(* IEC 61131-3 sources: POMIRTS_lab3/AS/Library_2/AsHydCon/V3.10.0 (part 2) *)

(* ---- AsHydCon.fun ---- *)
(********************************************************************
 * COPYRIGHT -- B&R
 ********************************************************************
 * Library: AsHydCon
 * File: AsHydCon.fun
 * Author: DI Thomas J. Frauscher
 * Created: July 2011
 ********************************************************************
 * Function blocks of library AsHydCon
 ********************************************************************)

FUNCTION_BLOCK HCRPT1 (*1st order delay element.*)
	VAR_INPUT
		enable : BOOL; (*Enable function block.*)
		V : REAL; (*Gain. Units: [1].*)
		T1 : REAL; (*Time constant. Units: [s]. Valid value range: T1 >= 0.*)
		u : REAL; (*Input value.*)
		Set_y : USINT; (*"Apply preset value for y" controller input. Valid value range: {0,1,2}.*)
		y_set : REAL; (*Preset value for y.*)
	END_VAR
	VAR_OUTPUT
		y : REAL; (*Output value.*)
		status : UINT; (*Function block status message.*)
	END_VAR
	VAR
		Internal : HCRPT1_Internal_typ; (*Data for internal use.*)
	END_VAR
END_FUNCTION_BLOCK

FUNCTION_BLOCK HCRPT2 (*2nd order delay element.*)
	VAR_INPUT
		enable : BOOL; (*Enable function block.*)
		V : REAL; (*Gain. Units: [1].*)
		T1 : REAL; (*Time constant 1. Units: [s]. Valid value range: T1 >= 0.*)
		T2 : REAL; (*Time constant 2. Units: [s]. Valid value range: T2 >= 0.*)
		u : REAL; (*Input value.*)
		Set_y : USINT; (*"Apply preset value for y" controller input. Valid value range: {0,1,2}.*)
		y_set : REAL; (*Preset value for y.*)
	END_VAR
	VAR_OUTPUT
		y : REAL; (*Output value.*)
		status : UINT; (*Function block status message.*)
	END_VAR
	VAR
		Internal : HCRPT2_Internal_typ; (*Data for internal use.*)
	END_VAR
END_FUNCTION_BLOCK

FUNCTION_BLOCK HCRPT2s (*Oscillating 2nd order delay element.*)
	VAR_INPUT
		enable : BOOL; (*Enable function block.*)
		V : REAL; (*Gain. Units: [1].*)
		D : REAL; (*Damping constant. Units: [1]. Valid value range: D >= 0.*)
		Tf : REAL; (*Filter time constant. Units: [s]. Valid value range: Tf > 0.*)
		u : REAL; (*Input value.*)
		Set_y : USINT; (*"Apply preset value for y" controller input. Valid value range: {0,1,2}.*)
		y_set : REAL; (*Preset value for y.*)
	END_VAR
	VAR_OUTPUT
		y : REAL; (*Output value.*)
		status : UINT; (*Function block status message.*)
	END_VAR
	VAR
		Internal : HCRPT2s_Internal_typ; (*Data for internal use.*)
	END_VAR
END_FUNCTION_BLOCK

FUNCTION_BLOCK HCRDT1 (*1st order differentiator.*)
	VAR_INPUT
		enable : BOOL; (*Enable function block.*)
		Tv : REAL; (*Differentiation time constant. Units: [s]. Valid value range: Tv >= 0.*)
		Tf : REAL; (*Filter time constant. Units: [s]. Valid value range: Tf >= 0.*)
		u : REAL; (*Input value.*)
		n_Avg : USINT; (*Moving average filter for the input value u. Valid value range: {0, 1, 2, ..., 100}.*)
		Reset_y : USINT; (*Reset controller input y to 0. Valid value range: {0,1,2}.*)
	END_VAR
	VAR_OUTPUT
		y : REAL; (*Output value.*)
		status : UINT; (*Function block status message.*)
	END_VAR
	VAR
		Internal : HCRDT1_Internal_typ; (*Data for internal use.*)
	END_VAR
END_FUNCTION_BLOCK

FUNCTION_BLOCK HCRDT2 (*2nd order differentiator.*)
	VAR_INPUT
		enable : BOOL; (*Enable function block.*)
		Tv : REAL; (*Differentiation time constant. Units: [s]. Valid value range: Tv >= 0.*)
		T1 : REAL; (*Filter time constant 1. Units: [s]. Valid value range: T1 >= 0.*)
		T2 : REAL; (*Filter time constant 2. Units: [s]. Valid value range: T2 >= 0.*)
		u : REAL; (*Input value.*)
		n_Avg : USINT; (*Moving average filter for the input value u. Valid value range: {0, 1, 2, ..., 100}.*)
		Reset_y : USINT; (*Reset controller input y to 0. Valid value range: {0,1,2}.*)
	END_VAR
	VAR_OUTPUT
		y : REAL; (*Output value.*)
		status : UINT; (*Function block status message.*)
	END_VAR
	VAR
		Internal : HCRDT2_Internal_typ; (*Data for internal use.*)
	END_VAR
END_FUNCTION_BLOCK

FUNCTION_BLOCK HCRDT2s (*Oscillating 2nd order differentiator.*)
	VAR_INPUT
		enable : BOOL; (*Enable function block.*)
		D : REAL; (*Damping constant. Units: [1]. Valid value range: D >= 0.*)
		Tv : REAL; (*Differentiation time constant. Units: [s]. Valid value range: Tv >= 0.*)
		Tf : REAL; (*Filter time constant. Units: [s]. Valid value range: Tf >= 0.*)
		u : REAL; (*Input value.*)
		Reset_y : USINT; (*Reset controller input y to 0. Valid value range: {0,1,2}.*)
	END_VAR
	VAR_OUTPUT
		y : REAL; (*Output value.*)
		status : UINT; (*Function block status message.*)
	END_VAR
	VAR
		Internal : HCRDT2s_Internal_typ; (*Data for internal use.*)
	END_VAR
END_FUNCTION_BLOCK

FUNCTION_BLOCK HCRIT1 (*1st order integrator.*)
	VAR_INPUT
		enable : BOOL; (*Enable function block.*)
		V : REAL; (*Gain. Units: [1].*)
		Tn : REAL; (*Integration time constant (integral action time). Units: [s]. Valid value range: Tn > 0.*)
		T1 : REAL; (*Time constant. Units: [s]. Valid value range: T1 >= 0.*)
		u : REAL; (*Input value.*)
		Set_y : USINT; (*"Apply preset value for y" controller input. Valid value range: {0,1,2}.*)
		y_set : REAL; (*Preset value for y.*)
	END_VAR
	VAR_OUTPUT
		y : REAL; (*Output value.*)
		status : UINT; (*Function block status message.*)
	END_VAR
	VAR
		Internal : HCRIT1_Internal_typ; (*Data for internal use.*)
	END_VAR
END_FUNCTION_BLOCK

FUNCTION_BLOCK HCRNotch (*2nd order notch filter.*)
	VAR_INPUT
		enable : BOOL; (*Enable function block.*)
		V : REAL; (*Gain. Units: [1].*)
		f0 : REAL; (*Filter frequency. Units: [Hz]. Valid value range: f0 > 0.*)
		B : REAL; (*Filter band width. Units: [Hz]. Valid value range: B > 0.*)
		u : REAL; (*Input value.*)
		Set_y : USINT; (*"Apply preset value for y" controller input. Valid value range: {0,1,2}.*)
		y_set : REAL; (*Preset value for y.*)
	END_VAR
	VAR_OUTPUT
		y : REAL; (*Output value.*)
		status : UINT; (*Function block status message.*)
	END_VAR
	VAR
		Internal : HCRNotch_Internal_typ; (*Data for internal use.*)
	END_VAR
END_FUNCTION_BLOCK

FUNCTION_BLOCK HCRPT1cP (*Converging 1st order delay element.*)
	VAR_INPUT
		enable : BOOL; (*Enable function block.*)
		T1 : REAL; (*Time constant. Units: [s]. Valid value range: T1 >= 0.*)
		u : REAL; (*Input value.*)
		Set_y : USINT; (*"Apply preset value for y" controller input. Valid value range: {0,1,2}.*)
		y_set : REAL; (*Preset value for y.*)
	END_VAR
	VAR_OUTPUT
		y : REAL; (*Output value.*)
		status : UINT; (*Function block status message.*)
	END_VAR
	VAR
		Internal : HCRPT1cP_Internal_typ; (*Data for internal use.*)
	END_VAR
END_FUNCTION_BLOCK

FUNCTION_BLOCK HCRJoltFree (*Jolt-free switching between 2 inputs.*)
	VAR_INPUT
		enable : BOOL; (*Enable function block.*)
		tSwitch : REAL; (*Switching time. Units: [s]. Valid value range: tSwitch >= 0.*)
		uSwitch : BOOL; (*Switch between signal inputs u1 and u2.*)
		u1 : REAL; (*Input value 1.*)
		u2 : REAL; (*Input value 2.*)
	END_VAR
	VAR_OUTPUT
		y : REAL; (*Output value.*)
		status : UINT; (*Function block status message.*)
	END_VAR
	VAR
		Internal : HCRJoltFree_Internal_typ; (*Data for internal use.*)
		PT1cP : HCRPT1cP; (*Internally used function block.*)
	END_VAR
END_FUNCTION_BLOCK

FUNCTION_BLOCK HCRFIFO (*FIFO (dead time) element.*)
	VAR_INPUT
		enable : BOOL; (*Enable function block.*)
		t_FIFO : DINT; (*Delay time. Units: [µs].*)
		x : REAL; (*Input value.*)
		Set_y : BOOL; (*"Apply preset value for y" controller input.*)
		y_set : REAL; (*Preset value for y.*)
	END_VAR
	VAR_OUTPUT
		y : REAL; (*Output value.*)
		status : UINT; (*Function block status message.*)
	END_VAR
	VAR
		Internal : HCRFIFO_Internal_typ; (*Data for internal use.*)
	END_VAR
END_FUNCTION_BLOCK

FUNCTION_BLOCK HCRRampGen (*Ramp generator.*)
	VAR_INPUT
		enable : BOOL; (*Enable function block.*)
		t_rise : REAL; (*Rise time. Units [s]. Valid value range: t_rise >= 0.*)
		t_hold : REAL; (*Constant holding time. Units [s]. Valid value range: t_hold >= 0.*)
		t_fall : REAL; (*Fall time. Units [s]. Valid value range: t_fall >= 0.*)
		y_start : REAL; (*Start value for the output value y.*)
		y_hold : REAL; (*Stop value for the output value y.*)
		y_end : REAL; (*End value for the output value y.*)
		Init : BOOL; (*Based on the start value y_start, Init = 1 initiates a new ramp that ends with an end value y_end, after crossing a stop phase t_hold with stop value y_hold.*)
	END_VAR
	VAR_OUTPUT
		y : REAL; (*Ramp generator output value.*)
		dy : REAL; (*Time derivative (dy/dt) of y.*)
		dy_ramped : REAL; (*Ramped time derivative (dy/dt) of y.*)
		Finished : BOOL; (*Finished = 1 indicates the end of ramp generation.*)
		status : UINT; (*Function block status message.*)
	END_VAR
	VAR
		Internal : HCRRampGen_Internal_typ; (*Data for internal use.*)
	END_VAR
END_FUNCTION_BLOCK

FUNCTION_BLOCK HCRSPF (*Smart path finder.*)
	VAR_INPUT
		enable : BOOL; (*Enable function block.*)
		pMove_Para : REFERENCE TO HCRMovePara_typ; (*Movement parameters (t_Jolt, vC_pos, vC_neg, aAcc_pos, aDec_pos, aAcc_neg, aDec_neg).*)
		Stop : BOOL; (*Stop = 1 stops trajectory planning.*)
		s_home : REAL; (*Homing position. Units: [mm].*)
		Set_home : BOOL; (*If no set trajectory is being processed at the moment, setting Set_home = 1 sets s_set = s_home and Reached = 1.*)
		s_end : REAL; (*End position of the trajectory. Units: [mm].*)
		Init : BOOL; (*Based on the current set position s_set and the current set speed v_set, Init = 1 initiates a new trajectory that ends at the point s_end.*)
		Brake : BOOL; (*Based on the current values of s_set and v_set, Brake = 1 stops the movement with the delay aDec_pos (positive direction) or aDec_neg (negative direction).*)
	END_VAR
	VAR_OUTPUT
		s_set : REAL; (*Set position. Units: [mm].*)
		v_set : REAL; (*Set speed. Units: [mm/s]. Value range: -vC_neg <= v_set <= vC_pos.*)
		a_set : REAL; (*Set acceleration. Units: [mm/s²]. Value range: -max(aDec_pos, aDec_neg) <= a_set <= max(aAcc_pos, aAcc_neg).*)
		MoveDir : SINT; (*Direction of movement. Value range: {-3,-2,-1: negative direction of movement (-3: Deceleration phase, -2: Constant speed phase, -1: Acceleration phase), 0: standstill, 1,2,3: positive direction of movement (1: Acceleration phase, 2: Constant speed phase, 3: Deceleration phase)}.*)
		ApproachDir : SINT; (*Approach direction indicates in which direction the end position s_end is reached. Value range: {-1: negative approach direction, 0: undefined, 1: positive approach direction}.*)
		Reached : BOOL; (*Reached = 1 indicates that the end position has been reached and that the movement is complete.*)
		status : UINT; (*Function block status message.*)
	END_VAR
	VAR
		Internal : HCRSPF_Internal_typ; (*Data for internal use.*)
		SystemInfo : SysInfo; (*Internally used function block.*)
	END_VAR
END_FUNCTION_BLOCK

FUNCTION_BLOCK HCRSFG (*Smart force generator.*)
	VAR_INPUT
		enable : BOOL; (*Enable function block.*)
		t_Jolt : REAL; (*Jolt time. Units [s]. Valid value range: 0 <= t_Jolt <= 0.2.*)
		Stop : BOOL; (*Stop = 1 stops trajectory planning.*)
		dFp_home : REAL; (*Homing value for the set force rate. Units: [N/s].*)
		Fp_home : REAL; (*Homing value for the set force. Units: [N].*)
		Set_home : BOOL; (*If no set trajectory is being processed at the moment, setting Set_home = 1 sets Fp_set = Fp_home, dFp_set = dFp_home and Reached = 1.*)
		t_delta : REAL; (*Time difference specified for bringing Fp_set from its present value to the end value Fp_end. Units: [s]. Valid value range: t_delta > t_Jolt.*)
		Fp_end : REAL; (*End value of the set force trajectory. Units: [N].*)
		Init : BOOL; (*Based on the current set force Fp_set and the current set force rate dFp_set, Init = 1 initiates a new trajectory that ends at the point Fp_end (dFp_set = 0).*)
	END_VAR
	VAR_OUTPUT
		Fp_set : REAL; (*Set force. Units: [N].*)
		dFp_set : REAL; (*Set force rate. Units: [N/s].*)
		t_delta_act : REAL; (*Actual time difference needed for bringing Fp_set to the specified end value Fp_end. Units: [s]. Value range: t_delta_act > t_Jolt.*)
		Reached : BOOL; (*Reached = 1 indicates that end value of the set force has been reached and that the profile generation is complete.*)
		status : UINT; (*Function block status message.*)
	END_VAR
	VAR
		Internal : HCRSFG_Internal_typ; (*Data for internal use.*)
		SPF : HCRSPF; (*Internally used function block.*)
	END_VAR
END_FUNCTION_BLOCK

FUNCTION_BLOCK HCRAutoTune (*Autotuning-algorithm for Kp.*)
	VAR_INPUT
		enable : BOOL; (*Enable function block.*)
		pSupply_max : REAL; (*Maximum system pressure (supply pressure). Units: [bar]. Valid value range: pSupply_max >= 0.*)
		A_Cyl_pos : REAL; (*Cylinder piston area whose pressurization induces a movement in the positive direction (e.g. extending piston). Units: [cm]. Valid value range: A_Cyl_pos > 0.*)
		A_Cyl_neg : REAL; (*Cylinder piston area whose pressurization induces a movement in the negative direction (e.g. retracting piston). Units: [cm]. Valid value range: A_Cyl_neg > 0.*)
		Qnom_pos : REAL; (*Nominal valve-volume flow, which, together with A_Cyl_pos results in a movement in the positive direction (e.g. extending piston). Units: [l/min]. Valid value range: Qnom_pos > 0.*)
		Qnom_neg : REAL; (*Nominal valve-volume flow, which, together with A_Cyl_neg results in a movement in the negative direction (e.g. retracting piston). Units: [l/min]. Valid value range: Qnom_neg > 0.*)
		pDelta_nom : REAL; (*Nominal pressure drop at valve edge. Units: [bar]. Valid value range: pDelta_nom > 0.*)
		V0_pos : REAL; (*Static volume in reference to the cylinder chamber responsible for movement in the 'positive' direction (e.g. extending piston). Units: [l]. Valid value range: V0_pos >= 0.*)
		V0_neg : REAL; (*Static volume in reference to the cylinder chamber responsible for movement in the 'negative' direction (e.g. retracting piston). Units: [l]. Valid value range: V0_neg >= 0.*)
		h_Cyl : REAL; (*Cylinder height. Units: [mm]. Valid value range: h_Cyl > 0.*)
		m_Cyl : REAL; (*Resulting mass of the moving hydraulic system. Units: [kg]. Valid value range: m_Cyl > 0.*)
		s_min : REAL; (*Minimum value of set position and actual position. Units: [mm]. Valid value range: s_min < s_max.*)
		s_max : REAL; (*Maximum value of set position and actual position. Units: [mm]. Valid value range: s_max > s_min.*)
		Update : USINT; (*Any changes to the above variables (pSupply_max, A_Cyl_pos, ..., s_max) must be applied with Update = 1.*)
	END_VAR
	VAR_OUTPUT
		Kp : REAL; (*Calculated proportional gain of the position controller. Units: [1].*)
		status : UINT; (*Function block status message.*)
	END_VAR
	VAR
		Internal : HCRAutoTune_Internal_typ; (*Data for internal use.*)
	END_VAR
END_FUNCTION_BLOCK

FUNCTION_BLOCK HCROmega0 (*Omega0-correction for Kp.*)
	VAR_INPUT
		enable : BOOL; (*Enable function block.*)
		A_Cyl_pos : REAL; (*Cylinder piston area whose pressurization induces a movement in the positive direction (e.g. extending piston). Units: [cm]. Valid value range: A_Cyl_pos > 0.*)
		A_Cyl_neg : REAL; (*Cylinder piston area whose pressurization induces a movement in the negative direction (e.g. retracting piston). Units: [cm]. Valid value range: A_Cyl_neg > 0.*)
		V0_pos : REAL; (*Static volume in reference to the cylinder chamber responsible for movement in the 'positive' direction (e.g. extending piston). Units: [l]. Valid value range: V0_pos >= 0.*)
		V0_neg : REAL; (*Static volume in reference to the cylinder chamber responsible for movement in the 'negative' direction (e.g. retracting piston). Units: [l]. Valid value range: V0_neg >= 0.*)
		h_Cyl : REAL; (*Cylinder height. Units: [mm]. Valid value range: h_Cyl > 0.*)
		x_Cyl_min : REAL; (*Minimum value of x_Cyl until a correction of the proportional gain of the position controller has been calculated. Units: [mm]. Valid value range: 0 <= x_Cyl_min < x_Cyl_max.*)
		x_Cyl_max : REAL; (*Maximum value of x_Cyl until a correction of the proportional gain of the position controller has been calculated. Units: [mm]. Valid value range: x_Cyl_min < x_Cyl_max <= h_Cyl.*)
		Update : USINT; (*Any changes to the above variables (A_Cyl_pos, A_Cyl_neg, ..., x_Cyl_max) must be applied with Update = 1.*)
		x_Cyl : REAL; (*Current position of the cylinder piston (always based on the cylinder). Units: [mm]. Valid value range: 0 <= x_Cyl <= h_Cyl.*)
	END_VAR
	VAR_OUTPUT
		x0_Cyl : REAL; (*Position of cylinder piston at which the critical natural frequency of the hydraulic system occurs. Units: [mm]. Value range: 0 <= x0_Cyl <= h_Cyl.*)
		Kp_xCorr : REAL; (*Calculated multiplication factor for correcting the proportional gain of the position controller with Kp_xCorr = Kp_xCorr(x_Cyl). Units: [1]. Value range: 1 <= Kp_xCorr <= 2.*)
		status : UINT; (*Function block status message.*)
	END_VAR
	VAR
		Internal : HCROmega0_Internal_typ; (*Data for internal use.*)
	END_VAR
END_FUNCTION_BLOCK

FUNCTION_BLOCK HCRvyServo (*v-y servo correction (pressure).*)
	VAR_INPUT
		enable : BOOL; (*Enable function block.*)
		pSupply_max : REAL; (*Maximum system pressure (supply pressure). Units: [bar]. Valid value range: pSupply_max >= 0.*)
		pSupply : REAL; (*System pressure (supply pressure). Units: [bar]. Valid value range: pSupply > 0.*)
		pTank : REAL; (*Tank pressure. Units: [bar]. Valid value range: pTank >= 0.*)
		A_Cyl_pos : REAL; (*Cylinder piston area whose pressurization induces a movement in the positive direction (e.g. extending piston). Units: [cm]. Valid value range: A_Cyl_pos > 0.*)
		A_Cyl_neg : REAL; (*Cylinder piston area whose pressurization induces a movement in the negative direction (e.g. retracting piston). Units: [cm]. Valid value range: A_Cyl_neg > 0.*)
		Qnom_pos : REAL; (*Nominal valve-volume flow, which, together with A_Cyl_pos results in a movement in the positive direction (e.g. extending piston). Units: [l/min]. Valid value range: Qnom_pos > 0.*)
		Qnom_neg : REAL; (*Nominal valve-volume flow, which, together with A_Cyl_neg results in a movement in the negative direction (e.g. retracting piston). Units: [l/min]. Valid value range: Qnom_neg > 0.*)
		pDelta_nom : REAL; (*Nominal pressure drop at valve edge. Units: [bar]. Valid value range: pDelta_nom > 0.*)
		yValve_0 : REAL; (*Valve overlap. Units: [1]. Valid value range:  0 <= yValve_0 < 1.*)
		yValve_min : REAL; (*Minimum valve opening (|yValve| = yValve_min). Units: [1]. Valid value range: 0 <= yValve_min <= 1.*)
		Neg_y : BOOL; (*Negative values for the valve opening yValve result in a positive speed, and vice versa (inverted valve behavior).*)
		Update : USINT; (*Any changes to the above variables must be applied with Update = (Mode + 1).*)
		pCyl_pos : REAL; (*Chamber pressure for movement in the 'positive' direction. Units: [bar]. Valid value range: 0 <= pCyl_pos < pSupply.*)
		pCyl_neg : REAL; (*Chamber pressure for movement in the 'negative' direction. Units: [bar]. Valid value range: 0 <= pCyl_neg < pSupply.*)
		vCyl_abs : REAL; (*Absolute speed of cylinder movement. Units: [mm/s]. Valid value range: -vCyl_sup < vCyl_abs < vCyl_sup.*)
		vCyl_rel : REAL; (*Relative speed of cylinder movement. Units: [%]. Valid value range: -100 <= vCyl_rel <= 100.*)
		Zero_yValve : BOOL; (*Setting this input results in the immediate output of yValve = 0 and Qy = 0.*)
	END_VAR
	VAR_OUTPUT
		Qy_abs : REAL; (*Volume flow produced by vCyl_abs (Qy = Qy_abs + Qy_rel). Units: [l/min]. Value range: -Qnom_neg <= Qy_abs <= Qnom_pos.*)
		Qy_rel : REAL; (*Volume flow produced by vCyl_rel (Qy_rel = Qy - Qy_abs). Units: [l/min]. Value range: -Qnom_neg <= Qy_rel <= Qnom_pos.*)
		Qy : REAL; (*Volume flow produced by valve opening yValve. Units: [l/min]. Value range: -Qnom_neg <= Qy <= Qnom_pos.*)
		yValve : REAL; (*Valve opening. Units: [1]. Value range: -1 <= yValve <= 1.*)
		MoveDir : SINT; (*Direction of movement. Value range: {-1: negative direction of movement, 0: undefined, 1: positive direction of movement}.*)
		status : UINT; (*Function block status message.*)
	END_VAR
	VAR
		Internal : HCRvyServo_Internal_typ; (*Data for internal use.*)
	END_VAR
END_FUNCTION_BLOCK

FUNCTION_BLOCK HCRvyServo_Fp (*v-y servo correction (force).*)
	VAR_INPUT
		enable : BOOL; (*Enable function block.*)
		pSupply_max : REAL; (*Maximum system pressure (supply pressure). Units: [bar]. Valid value range: pSupply_max >= 0.*)
		pSupply : REAL; (*System pressure (supply pressure). Units: [bar]. Valid value range: pSupply > 0.*)
		pTank : REAL; (*Tank pressure. Units: [bar]. Valid value range: pTank >= 0.*)
		A_Cyl_pos : REAL; (*Cylinder piston area whose pressurization induces a movement in the positive direction (e.g. extending piston). Units: [cm]. Valid value range: A_Cyl_pos > 0.*)
		A_Cyl_neg : REAL; (*Cylinder piston area whose pressurization induces a movement in the negative direction (e.g. retracting piston). Units: [cm]. Valid value range: A_Cyl_neg > 0.*)
		Qnom_pos : REAL; (*Nominal valve-volume flow, which, together with A_Cyl_pos results in a movement in the positive direction (e.g. extending piston). Units: [l/min]. Valid value range: Qnom_pos > 0.*)
		Qnom_neg : REAL; (*Nominal valve-volume flow, which, together with A_Cyl_neg results in a movement in the negative direction (e.g. retracting piston). Units: [l/min]. Valid value range: Qnom_neg > 0.*)
		pDelta_nom : REAL; (*Nominal pressure drop at valve edge. Units: [bar]. Valid value range: pDelta_nom > 0.*)
		yValve_0 : REAL; (*Valve overlap. Units: [1]. Valid value range:  0 <= yValve_0 < 1.*)
		yValve_min : REAL; (*Minimum valve opening (|yValve| = yValve_min). Units: [1]. Valid value range: 0 <= yValve_min <= 1.*)
		Neg_y : BOOL; (*Negative values for the valve opening yValve result in a positive speed, and vice versa (inverted valve behavior).*)
		Update : USINT; (*Any changes to the above variables must be applied with Update = (Mode + 1).*)
		Fp_Cyl : REAL; (*Process force. Units: [N].*)
		Ff_Cyl_pos : REAL; (*Friction force in positive direction. Units: [N]. Valid value range:  Ff_Cyl_pos >= 0.*)
		Ff_Cyl_neg : REAL; (*Friction force in negative direction. Units: [N]. Valid value range:  Ff_Cyl_neg >= 0.*)
		vCyl_abs : REAL; (*Absolute speed of cylinder movement. Units: [mm/s]. Valid value range: -vCyl_sup < vCyl_abs < vCyl_sup.*)
		vCyl_rel : REAL; (*Relative speed of cylinder movement. Units: [%]. Valid value range: -100 <= vCyl_rel <= 100.*)
		Zero_yValve : BOOL; (*Setting this input results in the immediate output of yValve = 0 and Qy = 0.*)
	END_VAR
	VAR_OUTPUT
		Qy_abs : REAL; (*Volume flow produced by vCyl_abs (Qy = Qy_abs + Qy_rel). Units: [l/min]. Value range: -Qnom_neg <= Qy_abs <= Qnom_pos.*)
		Qy_rel : REAL; (*Volume flow produced by vCyl_rel (Qy_rel = Qy - Qy_abs). Units: [l/min]. Value range: -Qnom_neg <= Qy_rel <= Qnom_pos.*)
		Qy : REAL; (*Volume flow produced by valve opening yValve. Units: [l/min]. Value range: -Qnom_neg <= Qy <= Qnom_pos.*)
		yValve : REAL; (*Valve opening. Units: [1]. Value range: -1 <= yValve <= 1.*)
		MoveDir : SINT; (*Direction of movement. Value range: {-1: negative direction of movement, 0: undefined, 1: positive direction of movement}.*)
		status : UINT; (*Function block status message.*)
	END_VAR
	VAR
		Internal : HCRvyServo_Fp_Internal_typ; (*Data for internal use.*)
	END_VAR
END_FUNCTION_BLOCK

FUNCTION_BLOCK HCRFyServo (*F-y servo correction (pressure).*)
	VAR_INPUT
		enable : BOOL; (*Enable function block.*)
		pSupply_max : REAL; (*Maximum system pressure (supply pressure). Units: [bar]. Valid value range: pSupply_max >= 0.*)
		pSupply : REAL; (*System pressure (supply pressure). Units: [bar]. Valid value range: pSupply > 0.*)
		pTank : REAL; (*Tank pressure. Units: [bar]. Valid value range: pTank >= 0.*)
		A_Cyl_pos : REAL; (*Cylinder piston area whose pressurization induces a movement in the positive direction (e.g. extending piston). Units: [cm]. Valid value range: A_Cyl_pos > 0.*)
		A_Cyl_neg : REAL; (*Cylinder piston area whose pressurization induces a movement in the negative direction (e.g. retracting piston). Units: [cm]. Valid value range: A_Cyl_neg > 0.*)
		Qnom_pos : REAL; (*Nominal valve-volume flow, which, together with A_Cyl_pos results in a movement in the positive direction (e.g. extending piston). Units: [l/min]. Valid value range: Qnom_pos > 0.*)
		Qnom_neg : REAL; (*Nominal valve-volume flow, which, together with A_Cyl_neg results in a movement in the negative direction (e.g. retracting piston). Units: [l/min]. Valid value range: Qnom_neg > 0.*)
		pDelta_nom : REAL; (*Nominal pressure drop at valve edge. Units: [bar]. Valid value range: pDelta_nom > 0.*)
		yValve_0 : REAL; (*Valve overlap. Units: [1]. Valid value range:  0 <= yValve_0 < 1.*)
		V0_pos : REAL; (*Static volume in reference to the cylinder chamber responsible for movement in the 'positive' direction (e.g. extending piston). Units: [l]. Valid value range: V0_pos >= 0.*)
		V0_neg : REAL; (*Static volume in reference to the cylinder chamber responsible for movement in the 'negative' direction (e.g. retracting piston). Units: [l]. Valid value range: V0_neg >= 0.*)
		h_Cyl : REAL; (*Cylinder height. Units: [mm]. Valid value range: h_Cyl > 0.*)
		Neg_y : BOOL; (*Negative values for the valve opening yValve result in a positive speed, and vice versa (inverted valve behavior).*)
		Update : USINT; (*Any changes to the above variables must be applied with Update = (Mode + 1).*)
		x_Cyl : REAL; (*Current position of the cylinder piston (always based on the cylinder). Units: [mm]. Valid value range: 0 <= x_Cyl <= h_Cyl.*)
		v_Cyl : REAL; (*Current speed of the cylinder piston (always based on the cylinder). Units: [mm].*)
		pCyl_pos : REAL; (*Chamber pressure for movement in the 'positive' direction. Units: [bar]. Valid value range: 0 <= pCyl_pos < pSupply.*)
		pCyl_neg : REAL; (*Chamber pressure for movement in the 'negative' direction. Units: [bar]. Valid value range: 0 <= pCyl_neg < pSupply.*)
		dF_Cyl_abs : REAL; (*Absolute rate of force increase of the cylinder. Units: [N/s]. Valid value range:  -dF_Cyl_sup < dF_Cyl_abs < dF_Cyl_sup.*)
		dF_Cyl_rel : REAL; (*Relative rate of force increase of the cylinder. Units: [%]. Valid value range: -100 <= dF_Cyl_rel <= 100.*)
	END_VAR
	VAR_OUTPUT
		Qy : REAL; (*Volume flow produced by valve opening yValve. Units: [l/min]. Value range: -Qnom_neg <= Qy <= Qnom_pos.*)
		yValve : REAL; (*Valve opening. Units: [1]. Value range: -1 <= yValve <= 1.*)
		status : UINT; (*Function block status message.*)
	END_VAR
	VAR
		Internal : HCRFyServo_Internal_typ; (*Data for internal use.*)
	END_VAR
END_FUNCTION_BLOCK

FUNCTION_BLOCK HCRFyServo_Fp (*F-y servo correction (force).*)
	VAR_INPUT
		enable : BOOL; (*Enable function block.*)
		pSupply_max : REAL; (*Maximum system pressure (supply pressure). Units: [bar]. Valid value range: pSupply_max >= 0.*)
		pSupply : REAL; (*System pressure (supply pressure). Units: [bar]. Valid value range: pSupply > 0.*)
		pTank : REAL; (*Tank pressure. Units: [bar]. Valid value range: pTank >= 0.*)
		A_Cyl_pos : REAL; (*Cylinder piston area whose pressurization induces a movement in the positive direction (e.g. extending piston). Units: [cm]. Valid value range: A_Cyl_pos > 0.*)
		A_Cyl_neg : REAL; (*Cylinder piston area whose pressurization induces a movement in the negative direction (e.g. retracting piston). Units: [cm]. Valid value range: A_Cyl_neg > 0.*)
		Qnom_pos : REAL; (*Nominal valve-volume flow, which, together with A_Cyl_pos results in a movement in the positive direction (e.g. extending piston). Units: [l/min]. Valid value range: Qnom_pos > 0.*)
		Qnom_neg : REAL; (*Nominal valve-volume flow, which, together with A_Cyl_neg results in a movement in the negative direction (e.g. retracting piston). Units: [l/min]. Valid value range: Qnom_neg > 0.*)
		yValve_0 : REAL; (*Valve overlap. Units: [1]. Valid value range:  0 <= yValve_0 < 1.*)
		Neg_y : BOOL; (*Negative values for the valve opening yValve result in a positive speed, and vice versa (inverted valve behavior).*)
		Update : USINT; (*Any changes to the above variables must be applied with Update = (Mode + 1).*)
		Fp : REAL; (*Process force. Units: [N].*)
		u : REAL; (*Input value. Units: [1]. Valid value range: -1 <= u <= 1.*)
	END_VAR
	VAR_OUTPUT
		Qy : REAL; (*Volume flow produced by valve opening yValve. Units: [l/min]. Value range: -Qnom_neg <= Qy <= Qnom_pos.*)
		yValve : REAL; (*Valve opening. Units: [1]. Value range: -1 <= yValve <= 1.*)
		status : UINT; (*Function block status message.*)
	END_VAR
	VAR
		Internal : HCRFyServo_Fp_Internal_typ; (*Data for internal use.*)
	END_VAR
END_FUNCTION_BLOCK

FUNCTION_BLOCK HCRLinSpline (*Linear spline function.*)
	VAR_INPUT
		enable : BOOL; (*Enable function block.*)
		NbNodes : UINT; (*Number of nodes from the node vector that are used to define the point-to-point linear function 'f(x)'. Valid value range: NbNodes >= 0.*)
		pNodeVec : REFERENCE TO HCRNode_typ; (*Pointer to the first node vector element to be used, which represents the basis of 'f(x)' ([(X1,Y1), (X2,Y2), ..., (Xn,Yn)]) and 'f-1(x)' ([(Y1,X1), (Y2,X2), ..., (Yn,Xn)]), and which is formed as an array of HCRNode_typ elements.*)
		Invert : BOOL; (*Invert = 1 inverts the point-to-point linear function 'f(x)'. Also, y = 'f-1(x)', which is based on the inverted node vector [(Y1,X1), (Y2,X2), ..., (Yn,Xn)].*)
		Smooth : USINT; (*Smoothing in the area of around the node (Xi,Yi) of 'f(x)' and (Yi,Xi) of 'f-1(x)'. Valid value range: {0: off, 1: on}.*)
		Rness : REAL; (*Smoothing factor. Valid value range: 0 <= Rness <= 1000.*)
		Update : BOOL; (*Any changes to the above variables (NbNodes, ..., Rness) must be applied with Update = 1.*)
		DisMode : SINT; (*Processing discontinuities in 'f(x)' and 'f-1(x)'. Valid value range: {-1, 0, 1}.*)
		x : REAL; (*Abscissa value of 'f(x)' or 'f-1(x)'. Valid value range: X1 <= x <= Xn or Y1 <= x <= Yn.*)
	END_VAR
	VAR_OUTPUT
		y : REAL; (*Ordinate value of 'f(x)' or 'f-1(x)'.*)
		status : UINT; (*Function block status message.*)
	END_VAR
	VAR
		Internal : HCRLinSpline_Internal_typ; (*Data for internal use.*)
	END_VAR
END_FUNCTION_BLOCK

FUNCTION_BLOCK HCRLinValve (*Valve linearization.*)
	VAR_INPUT
		enable : BOOL; (*Enable function block.*)
		NbNodes : UINT; (*Number of nodes from the node vector that are used to define the point-to-point linear valve characteristic curve linearization 'f-1(Q)'. Valid value range: NbNodes >= 0.*)
		pNodeVec : REFERENCE TO HCRNode_typ; (*Pointer to the node vector element that is to be used first, which is the basis for the valve characteristic curve 'f(U)' ([(U1,Q1), (U2,Q2), ..., (Un,Qn)]), and which consists of an array of HCRNode_typ elements.*)
		Neg_Qy : BOOL; (*Neg_Qy = 1 negates the valve volume flow Qy (abscissa value of 'f-1(Q)').*)
		Neg_Uy : BOOL; (*Neg_Uy = 1 negates the control voltage Uy of the valve, i.e. +10V is reduced to -10V.*)
		Update : BOOL; (*Any changes to the above variables (NbNodes, pNodeVec and Neg_Uy) must be applied with Update = 1.*)
		DisMode : SINT; (*Processing of discontinuities in 'f-1(Q)', as they occur in positive overlapped valves. Valid value range: {-1, 0, 1}.*)
		Qy : REAL; (*Nominal valve volume flow as abscissa value of 'f-1(Q)'. Units: [l/min]. Valid value range: Q1 <= Qy <= Qn.*)
	END_VAR
	VAR_OUTPUT
		Uy : REAL; (*Control voltage of the valve (Neg_Uy = 0: U1 <= Uy <= Un, Neg_Uy = 1: -Un <= Uy <= -U1). Units: [V].*)
		status : UINT; (*Function block status message.*)
	END_VAR
	VAR
		Internal : HCRLinValve_Internal_typ; (*Data for internal use.*)
		LinSpline : HCRLinSpline; (*Internally used function block.*)
	END_VAR
END_FUNCTION_BLOCK

FUNCTION_BLOCK HCRPID (*PID controller.*)
	VAR_INPUT
		enable : BOOL; (*Enable function block.*)
		Parameter : HCRPIDPara_typ; (*PID parameters.*)
		Update : USINT; (*Every change to the above PID parameter vector must be made active using Update = 1.*)
		W : REAL; (*Reference variable (set value). Valid value range: WX_min <= W  <= WX_max.*)
		X : REAL; (*Controlled variable (actual value). Valid value range: WX_min <= X  <= WX_max.*)
		Invert : BOOL; (*Inversion of the effective direction of the controller using Invert = 1.*)
		I_Switch : SINT; (*Switch for the I part. Valid value range: I_{-4, -3, -2, -1, 0, 1, 2, 3, 4}.*)
		CTRLmode : USINT; (*Controller operating mode. Valid value range: {0x00, 0x01, 0x02, 0x03, 0x04, 0x05, 0x06, 0x07, 0x08}.*)
		Yman : REAL; (*Manipulated variable for manual operation. Units: [%]. Valid value range: Y_min <= Yman <= Y_max.*)
		Yadd : REAL; (*Feed forward value. Units: [%]. Valid value range: -100 <= Yadd <= 100.*)
	END_VAR
	VAR_OUTPUT
		e : REAL; (*Control deviation (e = W - X). Value range: (WX_min - WX_max) <= e  <= (WX_max - WX_min).*)
		Yp : REAL; (*Proportional part. Units: [%]. Value range: -100 <= Yp <= 100.*)
		Yi : REAL; (*Integration part. Units: [%]. Value range: Y_min <= Yi <= Y_max.*)
		Yd : REAL; (*Differential part. Units: [%]. Value range: -100 <= Yd <= 100.*)
		Y : REAL; (*Manipulated variable. Unit: [%]. Value range: Y_min <= Y <= Y_max.*)
		status : UINT; (*Function block status message.*)
	END_VAR
	VAR
		Internal : HCRPID_Internal_typ; (*Data for internal use.*)
	END_VAR
END_FUNCTION_BLOCK

FUNCTION_BLOCK HCRP2P_Cont (*Point-to-point position controller.*)
	VAR_INPUT
		enable : BOOL; (*Enable function block.*)
		s_set : REAL; (*Set position. Units: [mm].*)
		s_act : REAL; (*Actual position. Units: [mm].*)
		Kp : REAL; (*Proportional gain. Units: [%/mm]. Valid value range: Kp > 0.*)
		P2Pmode : SINT; (*Operating mode - position controller. Valid value range: {-1, 0, 1}.*)
		pAddPar : REFERENCE TO HCRP2P_Cont_AddPar_typ; (*Additional control parameters and options (Y_P2P_min, Y_P2P_max, dY_max, Tn_pos, Tn_neg, I_Switch, Tv, Tf).*)
	END_VAR
	VAR_OUTPUT
		Y_P2P : REAL; (*Manipulated variable. Unit: [%]. Value range: -100 <= Y_P2P <= 100.*)
		Y_P2P_int : INT; (*Valve opening in integer format. Value range: -32760 <= Y_P2P_int <= 32760.*)
		status : UINT; (*Function block status message.*)
	END_VAR
	VAR
		Internal : HCRP2P_Cont_Internal_typ; (*Data for internal use.*)
		PID : HCRPID; (*Internally used function block.*)
	END_VAR
END_FUNCTION_BLOCK

FUNCTION_BLOCK HCRs_Cont (*Position controller (force).*)
	VAR_INPUT
		enable : BOOL; (*Enable function block.*)
		pSystem_Para : REFERENCE TO HCRSystemPara_typ; (*System parameter (pSupply_max, pSupply, pTank, A_Cyl_pos, A_Cyl_neg).*)
		pValve_Para : REFERENCE TO HCRValvePara_typ; (*Valve parameter (Qnom_pos, Qnom_neg, pDelta_nom, yValve_0, Neg_y).*)
		pPID_Para_s : REFERENCE TO HCRPIDPara_s_typ; (*PID parameter - position controller.*)
		vyServoMode : USINT; (*v-y servo correction mode. Valid value range: {0, 2, 4, 6, 8}.*)
		Update : USINT; (*Every change to vyServoMode or to the parameters of the above vectors must be made active using Update = 1.*)
		s_set : REAL; (*Set position. Units: [mm].*)
		s_act : REAL; (*Actual position. Units: [mm].*)
		Invert : BOOL; (*Inversion of the effective direction of the controller using Invert = 1.*)
		I_Switch : USINT; (*Switch for the I part of the PID. Valid value range: {0, 1, 2, 3, 4}.*)
		CTRLmode : USINT; (*Operating mode - position controller. Valid value range: {0x00, 0x01, 0x02, 0x03, 0x04, 0x05, 0x06, 0x07, 0x08}.*)
		v_man : REAL; (*Speed of movement in manual operation. Units: [mm/s]. Valid value range: v_min <= v_man <= v_max.*)
		v_add : REAL; (*Additional speed input. Units: [mm/s]. Valid value range: -vCyl_sup < v_add < vCyl_sup.*)
		v_set : REAL; (*Set speed for speed input control of the cylinder movement. Units: [mm/s]. Valid value range: -vCyl_sup < v_set < vCyl_sup.*)
		Fp_Cyl : REAL; (*Process force. Units: [N].*)
		Ff_Cyl_pos : REAL; (*Friction force in positive direction. Units: [N]. Valid value range:  Ff_Cyl_pos >= 0.*)
		Ff_Cyl_neg : REAL; (*Friction force in negative direction. Units: [N]. Valid value range:  Ff_Cyl_neg >= 0.*)
		Qy_Oset_ext : REAL; (*External volume flow offset. Units: [l/min].*)
		Oset_Mode : USINT; (*Selection switch for offset compensation. Valid value range: {00000000, ..., 01111111}.*)
	END_VAR
	VAR_OUTPUT
		Qy_s : REAL; (*Calculated volume flow. Units: [l/min]. Value range: -Qnom_neg <= Qy_s <= Qnom_pos.*)
		Qy_Oset_s : REAL; (*Additive volume flow for offset compensation. Units: [l/min].*)
		Qy : REAL; (*Volume flow. Units: [l/min]. Value range: -Qnom_neg <= Qy <= Qnom_pos.*)
		yValve : REAL; (*Valve opening. Units: [1]. Value range: -1 <= yValve <= 1.*)
		MoveDir : SINT; (*Direction of movement. Value range: {-1: negative direction of movement, 0: undefined, 1: positive direction of movement}.*)
		status : UINT; (*Function block status message.*)
	END_VAR
	VAR
		Internal : HCRs_Cont_Internal_typ; (*Data for internal use.*)
		PID : HCRPID; (*Internally used function block.*)
		vyServo_Fp : HCRvyServo_Fp; (*Internally used function block.*)
	END_VAR
END_FUNCTION_BLOCK

FUNCTION_BLOCK HCRs_Cont_p (*Position controller (pressure).*)
	VAR_INPUT
		enable : BOOL; (*Enable function block.*)
		pSystem_Para : REFERENCE TO HCRSystemPara_typ; (*System parameter (pSupply_max, pSupply, pTank, A_Cyl_pos, A_Cyl_neg).*)
		pValve_Para : REFERENCE TO HCRValvePara_typ; (*Valve parameter (Qnom_pos, Qnom_neg, pDelta_nom, yValve_0, Neg_y).*)
		pPID_Para_s : REFERENCE TO HCRPIDPara_s_typ; (*PID parameter - position controller.*)
		vyServoMode : USINT; (*v-y servo correction mode. Valid value range: {0, 2, 4, 6, 8}.*)
		Update : USINT; (*Every change to vyServoMode or to the parameters of the above vectors must be made active using Update = 1.*)
		s_set : REAL; (*Set position. Units: [mm].*)
		s_act : REAL; (*Actual position. Units: [mm].*)
		Invert : BOOL; (*Inversion of the effective direction of the controller using Invert = 1.*)
		I_Switch : USINT; (*Switch for the I part of the PID. Valid value range: {0, 1, 2, 3, 4}.*)
		CTRLmode : USINT; (*Operating mode - position controller. Valid value range: {0x00, 0x01, 0x02, 0x03, 0x04, 0x05, 0x06, 0x07, 0x08}.*)
		v_man : REAL; (*Speed of movement in manual operation. Units: [mm/s]. Valid value range: v_min <= v_man <= v_max.*)
		v_add : REAL; (*Additional speed input. Units: [mm/s]. Valid value range: -vCyl_sup < v_add < vCyl_sup.*)
		v_set : REAL; (*Set speed for speed input control of the cylinder movement. Units: [mm/s]. Valid value range: -vCyl_sup < v_set < vCyl_sup.*)
		pCyl_pos : REAL; (*Chamber pressure for movement in the 'positive' direction. Units: [bar]. Valid value range: 0 <= pCyl_pos < pSupply.*)
		pCyl_neg : REAL; (*Chamber pressure for movement in the 'negative' direction. Units: [bar]. Valid value range: 0 <= pCyl_neg < pSupply.*)
		Qy_Oset_ext : REAL; (*External volume flow offset. Units: [l/min].*)
		Oset_Mode : USINT; (*Selection switch for offset compensation. Valid value range: {00000000, ..., 01111111}.*)
	END_VAR
	VAR_OUTPUT
		Qy_s : REAL; (*Calculated volume flow. Units: [l/min]. Value range: -Qnom_neg <= Qy_s <= Qnom_pos.*)
		Qy_Oset_s : REAL; (*Additive volume flow for offset compensation. Units: [l/min].*)
		Qy : REAL; (*Volume flow. Units: [l/min]. Value range: -Qnom_neg <= Qy <= Qnom_pos.*)
		yValve : REAL; (*Valve opening. Units: [1]. Value range: -1 <= yValve <= 1.*)
		MoveDir : SINT; (*Direction of movement. Value range: {-1: negative direction of movement, 0: undefined, 1: positive direction of movement}.*)
		status : UINT; (*Function block status message.*)
	END_VAR
	VAR
		Internal : HCRs_Cont_p_Internal_typ; (*Data for internal use.*)
		PID : HCRPID; (*Internally used function block.*)
		vyServo : HCRvyServo; (*Internally used function block.*)
	END_VAR
END_FUNCTION_BLOCK

FUNCTION_BLOCK HCRF_Cont (*Force controller (force).*)
	VAR_INPUT
		enable : BOOL; (*Enable function block.*)
		pSystem_Para : REFERENCE TO HCRSystemPara_typ; (*System parameter (pSupply_max, pSupply, pTank, A_Cyl_pos, A_Cyl_neg).*)
		pValve_Para : REFERENCE TO HCRValvePara_typ; (*Valve parameter (Qnom_pos, Qnom_neg, pDelta_nom, yValve_0, Neg_y).*)
		pPID_Para_F : REFERENCE TO HCRPIDPara_F_typ; (*PID parameter - force controller.*)
		FyServoMode : USINT; (*F-y servo correction mode. Valid value range: {0, 2, 8}.*)
		Update : USINT; (*Every change to FyServoMode or to the parameters of the above vectors must be made active using Update = 1.*)
		Fp_set : REAL; (*Set force. Units: [N].*)
		Fp_act : REAL; (*Actual force. Units: [N].*)
		Invert : BOOL; (*Inversion of the effective direction of the controller using Invert = 1.*)
		I_Switch : USINT; (*Switch for the I part of the PID. Valid value range: {0, 1, 2, 3, 4}.*)
		CTRLmode : USINT; (*Operating mode - force controller. Valid value range: {0x00, 0x01, 0x02, 0x03, 0x04, 0x05, 0x06, 0x07, 0x08, 0x10, 0x20}.*)
		Q_man : REAL; (*Valve volume flow in manual operation. Units: [l/min]. Valid value range: -Q_min <= Q_man <= Q_max.*)
		Q_add : REAL; (*Additional volume flow input. Units: [l/min]. Valid value range: -Qnom_neg <= Q_add <= Qnom_pos.*)
		v_act : REAL; (*Actual speed of the cylinder piston. Units: [mm/s].*)
		Qy_Oset_ext : REAL; (*External volume flow offset. Units: [l/min].*)
		Oset_Mode : USINT; (*Selection switch for offset compensation. Valid value range: {00000000, ..., 01111111}.*)
	END_VAR
	VAR_OUTPUT
		Qy_F : REAL; (*Calculated volume flow. Units: [l/min]. Value range: -Qnom_neg <= Qy_F <= Qnom_pos.*)
		Qy_Oset_F : REAL; (*Additive volume flow for offset compensation. Units: [l/min].*)
		Qy : REAL; (*Volume flow. Units: [l/min]. Value range: -Qnom_neg <= Qy <= Qnom_pos.*)
		yValve : REAL; (*Valve opening. Units: [1]. Value range: -1 <= yValve <= 1.*)
		status : UINT; (*Function block status message.*)
	END_VAR
	VAR
		Internal : HCRF_Cont_Internal_typ; (*Data for internal use.*)
		PID : HCRPID; (*Internally used function block.*)
		FyServo_Fp : HCRFyServo_Fp; (*Internally used function block.*)
	END_VAR
END_FUNCTION_BLOCK

FUNCTION_BLOCK HCRF_Cont_p (*Force controller (pressure).*)
	VAR_INPUT
		enable : BOOL; (*Enable function block.*)
		pSystem_Para : REFERENCE TO HCRSystemPara_typ; (*System parameter (pSupply_max, pSupply, pTank, A_Cyl_pos, A_Cyl_neg).*)
		pSystem_ParaAdd : REFERENCE TO HCRSystemParaAdd_typ; (*Additional system parameter (V0_pos, V0_neg, h_Cyl, m_Cyl).*)
		pValve_Para : REFERENCE TO HCRValvePara_typ; (*Valve parameter (Qnom_pos, Qnom_neg, pDelta_nom, yValve_0, Neg_y).*)
		pPID_Para_F : REFERENCE TO HCRPIDPara_F_typ; (*PID parameter - force controller.*)
		FyServoMode : USINT; (*F-y servo correction mode. Valid value range: {0, 2, 8}.*)
		Update : USINT; (*Every change to FyServoMode or to the parameters of the above vectors must be made active using Update = 1.*)
		Fp_set : REAL; (*Set force. Units: [N].*)
		Fp_act : REAL; (*Actual force. Units: [N].*)
		Invert : BOOL; (*Inversion of the effective direction of the controller using Invert = 1.*)
		I_Switch : USINT; (*Switch for the I part of the PID. Valid value range: {0, 1, 2, 3, 4}.*)
		CTRLmode : USINT; (*Operating mode - force controller. Valid value range: {0x00, 0x01, 0x02, 0x03, 0x04, 0x05, 0x06, 0x07, 0x08, 0x30}.*)
		Q_man : REAL; (*Valve volume flow in manual operation. Units: [l/min]. Valid value range: -Q_min <= Q_man <= Q_max.*)
		Q_add : REAL; (*Additional volume flow input. Units: [l/min]. Valid value range: -Qnom_neg <= Q_add <= Qnom_pos.*)
		dFp_set : REAL; (*Set value of the rate of force increase of the cylinder. Units: [N/s].*)
		x_Cyl : REAL; (*Current position of the cylinder piston (always based on the cylinder). Units: [mm]. Valid value range: 0 <= x_Cyl <= h_Cyl.*)
		v_Cyl : REAL; (*Current speed of the cylinder piston (always based on the cylinder). Units: [mm/s].*)
		pCyl_pos : REAL; (*Chamber pressure for movement in the 'positive' direction. Units: [bar]. Valid value range: 0 <= pCyl_pos < pSupply.*)
		pCyl_neg : REAL; (*Chamber pressure for movement in the 'negative' direction. Units: [bar]. Valid value range: 0 <= pCyl_neg < pSupply.*)
		v_act : REAL; (*Actual speed of the cylinder piston. Units: [mm/s].*)
		Qy_Oset_ext : REAL; (*External volume flow offset. Units: [l/min].*)
		Oset_Mode : USINT; (*Selection switch for offset compensation. Valid value range: {00000000, ..., 01111111}.*)
	END_VAR
	VAR_OUTPUT
		Qy_F : REAL; (*Calculated volume flow. Units: [l/min]. Value range: -Qnom_neg <= Qy_F <= Qnom_pos.*)
		Qy_Oset_F : REAL; (*Additive volume flow for offset compensation. Units: [l/min].*)
		Qy : REAL; (*Volume flow. Units: [l/min]. Value range: -Qnom_neg <= Qy <= Qnom_pos.*)
		yValve : REAL; (*Valve opening. Units: [1]. Value range: -1 <= yValve <= 1.*)
		status : UINT; (*Function block status message.*)
	END_VAR
	VAR
		Internal : HCRF_Cont_p_Internal_typ; (*Data for internal use.*)
		PID : HCRPID; (*Internally used function block.*)
		FyServo : HCRFyServo; (*Internally used function block.*)
	END_VAR
END_FUNCTION_BLOCK

FUNCTION_BLOCK HCRsF_Cont (*Switchable position/force controller (force).*)
	VAR_INPUT
		enable : BOOL; (*Enable function block.*)
		pSystem_Para : REFERENCE TO HCRSystemPara_typ; (*System parameter (pSupply_max, pSupply, pTank, A_Cyl_pos, A_Cyl_neg).*)
		pValve_Para : REFERENCE TO HCRValvePara_typ; (*Valve parameter (Qnom_pos, Qnom_neg, pDelta_nom, yValve_0, Neg_y).*)
		pPID_Para_s : REFERENCE TO HCRPIDPara_s_typ; (*PID parameter - position controller.*)
		pPID_Para_F : REFERENCE TO HCRPIDPara_F_typ; (*PID parameter - force controller.*)
		vyServoMode : USINT; (*v-y servo correction mode. Valid value range: {0, 2, 4, 6, 8}.*)
		FyServoMode : USINT; (*F-y servo correction mode. Valid value range: {0, 2, 8}.*)
		tSwitch : REAL; (*Switching time. Units: [s]. Valid value range: tSwitch >= 0.*)
		Update : USINT; (*Every change to vyServoMode, FyServoMode and tSwitch or to the parameters of the above vectors must be made active using Update = 1.*)
		s_set : REAL; (*Set position. Units: [mm].*)
		s_act : REAL; (*Actual position. Units: [mm].*)
		s_Cont_InVar : HCRs_Cont_InVar_typ; (*Additional input values - position controller.*)
		Fp_set : REAL; (*Set force. Units: [N].*)
		Fp_act : REAL; (*Actual force. Units: [N].*)
		F_Cont_InVar : HCRF_Cont_InVar_typ; (*Additional input values - force controller.*)
		CTRLmode : USINT; (*Operating mode. Valid value range: {0x00, 0x01, 0x02, 0x03, 0x04, 0x05, 0x06, 0x07, 0x08, 0x10, 0x20}.*)
		uSwitch : USINT; (*Switches between position controller and force controller.*)
	END_VAR
	VAR_OUTPUT
		Qy_s : REAL; (*Calculated volume flow (position). Units: [l/min]. Value range: -Qnom_neg <= Qy_s <= Qnom_pos.*)
		Qy_Oset_s : REAL; (*Additive volume flow for offset compensation (position). Units: [l/min].*)
		Qy_F : REAL; (*Calculated volume flow (force). Units: [l/min]. Value range: -Qnom_neg <= Qy_F <= Qnom_pos.*)
		Qy_Oset_F : REAL; (*Additive volume flow for offset compensation (force). Units: [l/min].*)
		Qy : REAL; (*Volume flow. Units: [l/min]. Value range: -Qnom_neg <= Qy <= Qnom_pos.*)
		yValve : REAL; (*Valve opening. Units: [1]. Value range: -1 <= yValve <= 1.*)
		MoveDir : SINT; (*Direction of movement. Value range: {-1: negative direction of movement, 0: undefined, 1: positive direction of movement}.*)
		InForceCtrl : BOOL; (*Force controller active.*)
		status : UINT; (*Function block status message.*)
	END_VAR
	VAR
		Internal : HCRsF_Cont_Internal_typ; (*Data for internal use.*)
		s_Cont : HCRs_Cont; (*Internally used function block.*)
		F_Cont : HCRF_Cont; (*Internally used function block.*)
		JoltFree : HCRJoltFree; (*Internally used function block.*)
	END_VAR
END_FUNCTION_BLOCK

FUNCTION_BLOCK HCRsF_Cont_p (*Switchable position/force controller (pressure).*)
	VAR_INPUT
		enable : BOOL; (*Enable function block.*)
		pSystem_Para : REFERENCE TO HCRSystemPara_typ; (*System parameter (pSupply_max, pSupply, pTank, A_Cyl_pos, A_Cyl_neg).*)
		pSystem_ParaAdd : REFERENCE TO HCRSystemParaAdd_typ; (*Additional system parameter (V0_pos, V0_neg, h_Cyl, m_Cyl).*)
		pValve_Para : REFERENCE TO HCRValvePara_typ; (*Valve parameter (Qnom_pos, Qnom_neg, pDelta_nom, yValve_0, Neg_y).*)
		pPID_Para_s : REFERENCE TO HCRPIDPara_s_typ; (*PID parameter - position controller.*)
		pPID_Para_F : REFERENCE TO HCRPIDPara_F_typ; (*PID parameter - force controller.*)
		vyServoMode : USINT; (*v-y servo correction mode. Valid value range: {0, 2, 4, 6, 8}.*)
		FyServoMode : USINT; (*F-y servo correction mode. Valid value range: {0, 2, 8}.*)
		tSwitch : REAL; (*Switching time. Units: [s]. Valid value range: tSwitch >= 0.*)
		Update : USINT; (*Every change to vyServoMode, FyServoMode and tSwitch or to the parameters of the above vectors must be made active using Update = 1.*)
		s_set : REAL; (*Set position. Units: [mm].*)
		s_act : REAL; (*Actual position. Units: [mm].*)
		s_Cont_p_InVar : HCRs_Cont_p_InVar_typ; (*Additional input values - position controller.*)
		Fp_set : REAL; (*Set force. Units: [N].*)
		Fp_act : REAL; (*Actual force. Units: [N].*)
		F_Cont_InVar : HCRF_Cont_p_InVar_typ; (*Additional input values - force controller.*)
		CTRLmode : USINT; (*Operating mode. Valid value range: {0x00, 0x01, 0x02, 0x03, 0x04, 0x05, 0x06, 0x07, 0x08, 0x10, 0x20, 0x30}.*)
		uSwitch : USINT; (*Switches between position controller and force controller.*)
	END_VAR
	VAR_OUTPUT
		Qy_s : REAL; (*Calculated volume flow (position). Units: [l/min]. Value range: -Qnom_neg <= Qy_s <= Qnom_pos.*)
		Qy_Oset_s : REAL; (*Additive volume flow for offset compensation (position). Units: [l/min].*)
		Qy_F : REAL; (*Calculated volume flow (force). Units: [l/min]. Value range: -Qnom_neg <= Qy_F <= Qnom_pos.*)
		Qy_Oset_F : REAL; (*Additive volume flow for offset compensation (force). Units: [l/min].*)
		Qy : REAL; (*Volume flow. Units: [l/min]. Value range: -Qnom_neg <= Qy <= Qnom_pos.*)
		yValve : REAL; (*Valve opening. Units: [1]. Value range: -1 <= yValve <= 1.*)
		MoveDir : SINT; (*Direction of movement. Value range: {-1: negative direction of movement, 0: undefined, 1: positive direction of movement}.*)
		InForceCtrl : BOOL; (*Force controller active.*)
		status : UINT; (*Function block status message.*)
	END_VAR
	VAR
		Internal : HCRsF_Cont_p_Internal_typ; (*Data for internal use.*)
		s_Cont_p : HCRs_Cont_p; (*Internally used function block.*)
		F_Cont : HCRF_Cont; (*Internally used function block.*)
		F_Cont_p : HCRF_Cont_p; (*Internally used function block.*)
		vyServo : HCRvyServo; (*Internally used function block.*)
		JoltFree : HCRJoltFree; (*Internally used function block.*)
	END_VAR
END_FUNCTION_BLOCK

(* ---- AsHydCon.var ---- *)
(********************************************************************
 * COPYRIGHT -- B&R
 ********************************************************************
 * Library: AsHydCon
 * File: AsHydCon.var
 * Author: DI Thomas J. Frauscher
 * Created: July 2011
 ********************************************************************
 * Constants of library AsHydCon
 ********************************************************************)
VAR CONSTANT
  HCR_ERR_DT12S_D_NEG : UINT := 32250; (*Error: The damping constant D is negative.*)
  HCR_ERR_DT12S_T1_NEG : UINT := 32251; (*Error: The filter time constant T1 is negative.*)
  HCR_ERR_DT12S_T1_T2_ZERO : UINT := 32252; (*No longer used.*)
  HCR_ERR_DT12S_T2_NEG : UINT := 32253; (*Error: The filter time constant T2 is negative.*)
  HCR_ERR_DT12S_TF_NEG_ZERO : UINT := 32254; (*Error: The filter time constant Tf is less than or equal to 0.*)
  HCR_ERR_DT12S_TV_NEG : UINT := 32255; (*Error: The differentiation time constant Tv is negative.*)
  HCR_ERR_FIFO_MEM : UINT := 32256; (*Error: An error occurred during memory allocation for the internal ring buffer.*)
  HCR_ERR_FIFO_T_FIFO_NEG : UINT := 32257; (*Error: t_FIFO is negative.*)
  HCR_ERR_JFREE_TSWITCH_NEG : UINT := 32258; (*Error: The switching time tSwitch is negative.*)
  HCR_ERR_LIN_NODEVEC_EMPTY : UINT := 32259; (*Error: No valid pointer pNodeVec to the node vector found.*)
  HCR_ERR_LIN_X_NOT_ASC_DESC : UINT := 32260; (*Error: The x coordinates of the node vector are not sorted in ascending or descending order.*)
  HCR_ERR_LIN_Y_NOT_ASC_DESC : UINT := 32261; (*Error: The y coordinates (Ui with i = 1..n) of the node vector are not sorted in ascending or descending order.*)
  HCR_ERR_PID_DY_MAX_NEG : UINT := 32262; (*Error:
PID: The maximum manipulated variable ramp dY_max is negative.
Position controller: The maximum change rate for the piston speed (acceleration) dv_max is negative.
Force controller: The maximum volume flow change speed dQ_max is negative.*)
  HCR_ERR_PID_D_MODE_INVALID : UINT := 32263; (*Error: Invalid differentiation mode (d_mode).*)
  HCR_ERR_PID_KW_0_1 : UINT := 32264; (*Error: The set value weakening factor Kw is less than 0 or greater than 1.*)
  HCR_ERR_PID_K_FBK_NEG : UINT := 32265; (*Error: The wind-up damping factor K_Fbk is negative.*)
  HCR_ERR_PID_TF_NEG : UINT := 32266; (*Error: The filter time constant Tf of the differentiator is negative.*)
  HCR_ERR_PID_TF_ZERO : UINT := 32267; (*No longer used.*)
  HCR_ERR_PID_TN_NEG_NEG : UINT := 32268; (*Error:
PID: The integration time constant for I_Switch < 0 Tn_neg is negative.
Position controller: The integration time constant for movements in the 'negative' direction Tn_neg is negative.*)
  HCR_ERR_PID_TN_POS_NEG : UINT := 32269; (*Error:
PID: The integration time constant for I_Switch > 0 Tn_pos is negative.
Position controller: The integration time constant for movements in the 'positive' direction Tn_pos is negative.
Force controller: The integration time constant Tn is negative.*)
  HCR_ERR_PID_TV_NEG : UINT := 32270; (*Error: The differentiation time constant Tv of the differentiator is negative.*)
  HCR_ERR_PID_WX_MAX_MIN : UINT := 32271; (*Error:
PID: The maximum set and/or actual value WX_max is lower than the minimum value WX_min.
Position controller: The maximum value of the set and/or actual position s_max is lower than the minimum value s_min.
Force controller: The maximum value of the set and/or actual force Fp_max is lower than the minimum value Fp_min.*)
  HCR_ERR_PID_Y_MAX_MIN : UINT := 32272; (*Error:
PID: The lower limit for manipulated variables Y_min is less than -100%, the upper limit for manipulated variables Y_max is greater than +100%, or Y_max is less than or equal to Y_min.
Position controller, AutoTune: The lower limit for piston speed v_min is less than -Internal.vCyl_sup, the upper limit for piston speed v_max is greater than Internal.vCyl_sup, or v_max is less than or equal to v_min.
Force controller: The lower limit for the valve volume flow Q_min is less than -Qnom_neg, the upper limit for the valve volume flow Q_max is greater than Qnom_pos or Q_max is less than or equal to Q_min.*)
  HCR_ERR_PT12_T1_NEG : UINT := 32273; (*Error: The time constant T1 is negative.*)
  HCR_ERR_PT12_T2_NEG : UINT := 32274; (*Error: The time constant T2 is negative.*)
  HCR_ERR_PT1CP_T1_NEG : UINT := 32275; (*Error: The time constant T1 is negative.*)
  HCR_ERR_PT2S_D_NEG : UINT := 32276; (*Error: The damping constant D is negative.*)
  HCR_ERR_PT2S_TF_NEG_ZERO : UINT := 32277; (*Error: The filter time constant Tf is less than or equal to 0.*)
  HCR_ERR_SERVO_Y_MIN : UINT := 32278; (*Error: The value of minimum valve opening is outside the permissible range of 0 <= yValve_min <= 1.*)
  HCR_ERR_SYSTEM_A_CYL : UINT := 32279; (*Error: At least one of the two cylinder piston areas A_Cyl_pos or A_Cyl_neg was entered as less than or equal to 0.*)
  HCR_ERR_SYSTEM_P_DIFF : UINT := 32280; (*Error: The tank pressure pTank is above the system pressure pSupply.*)
  HCR_ERR_SYSTEM_P_SUPPLY : UINT := 32281; (*Error: The system pressure pSupply is less than or equal to 0.*)
  HCR_ERR_SYSTEM_P_TANK : UINT := 32282; (*Error: The tank pressure pTank is negative.*)
  HCR_ERR_VALVE_P_DELTA_NOM : UINT := 32283; (*Error: The nominal pressure drop at valve edge pDelta_nom is less than or equal to 0.*)
  HCR_ERR_VALVE_Q_NOM : UINT := 32284; (*Error: At least one nominal valve volume flow (Qnom_pos or Qnom_neg) was entered as less than or equal to 0.*)
  HCR_ERR_VALVE_Y_0 : UINT := 32285; (*Error: The value of valve overlap is outside the valid range of 0 <= yValve_0 < 1.*)
  HCR_ERR_RAMP_T_FALL_NEG : UINT := 32286; (*Error: The fall time t_fall is negative.*)
  HCR_ERR_RAMP_T_HOLD_NEG : UINT := 32287; (*Error: The hold time t_hold is negative.*)
  HCR_ERR_RAMP_T_RISE_NEG : UINT := 32288; (*Error: The rise time t_rise is negative.*)
  HCR_ERR_SPF_A_ACC_NEG_NEG_ZERO : UINT := 32289; (*Error: Acceleration in the 'negative' direction aAcc_neg is negative.*)
  HCR_ERR_SPF_A_ACC_POS_NEG_ZERO : UINT := 32290; (*Error: Acceleration in the 'positive' direction aAcc_pos is negative.*)
  HCR_ERR_SPF_A_DEC_NEG_NEG_ZERO : UINT := 32291; (*Error: Deceleration in the 'negative' direction aDec_neg is negative.*)
  HCR_ERR_SPF_A_DEC_POS_NEG_ZERO : UINT := 32292; (*Error: Deceleration in the 'positive' direction aDec_pos is negative.*)
  HCR_ERR_SPF_NIL_PTR : UINT := 32293; (*Error: The pointer pMove_Para on the motion parameter vector is an NIL-Pointer.*)
  HCR_ERR_SPF_T_JOLT_NEG : UINT := 32294; (*Error: The jolt time t_Jolt is negative.*)
  HCR_ERR_SPF_VC_NEG_NEG_ZERO : UINT := 32295; (*Error: The maximum speed of movement in the 'negative' direction vC_neg is negative.*)
  HCR_ERR_SPF_VC_POS_NEG_ZERO : UINT := 32296; (*Error: The maximum speed of movement in the 'positive' direction vC_pos is negative.*)
  HCR_ERR_SYSTEM_H_CYL : UINT := 32297; (*Error: The cylinder height was entered as less than or equal to 0.*)
  HCR_ERR_SYSTEM_M_CYL : UINT := 32298; (*Error: The resulting moving mass of the hydraulic system was set less than or equal to 0.*)
  HCR_ERR_SYSTEM_NIL_PTR : UINT := 32299; (*Error: No pointer pSystem_Para (pSystem_ParaAdd) specified for the system parameters HCRSystemPara_typ (HCRSystemParaAdd_typ).*)
  HCR_ERR_SYSTEM_P_SUPPLY_MAX : UINT := 32300; (*Error: The maximum system pressure pSupply_max is less than 0.*)
  HCR_ERR_SYSTEM_V0_NEG : UINT := 32301; (*Error: The static volume of the cylinder chamber responsible for movement in the'negative' direction was set less than 0.*)
  HCR_ERR_SYSTEM_V0_POS : UINT := 32302; (*Error: The static volume of the cylinder chamber responsible for movement in the 'positive' direction was set less than 0.*)
  HCR_ERR_SERVO_MODE_FY : UINT := 32303; (*Error: The selected mode for the F-y servo correction does not exist.*)
  HCR_ERR_SERVO_MODE_VY : UINT := 32304; (*Error: The selected mode for the v-y servo correction does not exist.*)
  HCR_ERR_PID_NIL_PTR : UINT := 32305; (*Error:
Position controller: No pointer pPID_Para_s specified for the PID-parameters HCRPIDPara_s_typ.
Force controller: No pointer pPID_Para_F specified for the PID-parameters HCRPIDPara_F_typ.*)
  HCR_ERR_VALVE_NIL_PTR : UINT := 32306; (*Error: No pointer pValve_Para specified for the valve parameters HCRValvePara_typ.*)
  HCR_ERR_NOTCH_B_NEG_ZERO : UINT := 32307; (*Error: The filter band width B is less than or equal to 0.*)
  HCR_ERR_NOTCH_F0_NEG_ZERO : UINT := 32308; (*Error: The filter frequency f0 is less than or equal to 0.*)
  HCR_ERR_OMEGA0_X0_CYL : UINT := 32309; (*Error: Position of cylinder piston x0_Cyl, at which the critical natural frequency of the hydraulic system occurs, lies outside the cylinder dimensions.*)
  HCR_ERR_OMEGA0_X_CYL_MIN_MAX : UINT := 32310; (*Error: The minimum cylinder piston position value, after which the proportional gain correction is calculated is less than 0. The maximum position value, up to which the proportional gain is calculated is greater than the cylinder height h_Cyl or x_Cyl_max is less than or equal to x_Cyl_min.*)
  HCR_ERR_IT1_T1_NEG : UINT := 32313; (*Error: The time constant T1 is negative.*)
  HCR_ERR_IT1_TN_NEG_ZERO : UINT := 32314; (*Error: The integration time constant Tn is less than or equal to 0.*)
  HCR_ERR_SFG_T_DELTA_NEG_ZERO : UINT := 32315; (*Error: The time t_delta, which is available for the profile generation, is less than or equal to 0.*)
  HCR_ERR_SFG_T_DIFF : UINT := 32316; (*Error: The net time (t_delta - t_Jolt), which is available for the profile generation, is less than or equal to 0.*)
  HCR_ERR_SFG_T_JOLT_NEG : UINT := 32317; (*Error: The jolt time t_Jolt is negative.*)
  HCR_ERR_DT12S_TF_NEG : UINT := 32318; (*Error: The filter time constant Tf is less than 0.*)
  HCR_WARN_DT12S_T1_TS : UINT := 32370; (*Warning: The filter time constant T1 entered is not larger than the corresponding task cycle time.*)
  HCR_WARN_DT12S_T1_ZERO : UINT := 32371; (*Warning: The filter time constant T1 = 0.*)
  HCR_WARN_DT12S_T2_TS : UINT := 32372; (*Warning: The filter time constant T2 entered is not larger than the corresponding task cycle time.*)
  HCR_WARN_DT12S_T2_ZERO : UINT := 32373; (*Warning: The filter time constant T2 = 0.*)
  HCR_WARN_DT12S_TF_TS : UINT := 32374; (*Warning: The filter time constant Tf entered is not larger than the corresponding task cycle time.*)
  HCR_WARN_DT12S_TV_TS : UINT := 32375; (*Warning: The differentiation time constant Tv entered is not larger than the corresponding task cycle time.*)
  HCR_WARN_DT12S_TV_ZERO : UINT := 32376; (*Warning: The differentiation time constant Tv = 0.*)
  HCR_WARN_FIFO_T_FIFO_INT : UINT := 32377; (*Warning: t_FIFO was not entered as a whole number multiple of the cycle time.*)
  HCR_WARN_FIFO_T_FIFO_TS : UINT := 32378; (*Warning: t_FIFO was entered as smaller than the corresponding task cycle time, and was automatically increased to this value.*)
  HCR_WARN_JFREE_TSWITCH_5TS : UINT := 32379; (*Warning: The switching time tSwitch entered is not 5 times larger than the corresponding task cycle time.*)
  HCR_WARN_JFREE_TSWITCH_ZERO : UINT := 32380; (*Warning: The switching time tSwitch = 0.*)
  HCR_WARN_LIN_CRIT_RNESS : UINT := 32381; (*Warning: The smoothing factor Rness is larger than the maximum possible smoothing factor (Internal.Rness_crit).*)
  HCR_WARN_LIN_NB_NODE : UINT := 32382; (*Warning: NbNodes <= 1.*)
  HCR_WARN_LIN_X_NOT_ASC_DESC_S : UINT := 32383; (*Warning: Sorting of the x coordinates of the node vector is monotonic, but not strictly monotonic.*)
  HCR_WARN_LIN_Y_NOT_ASC_DESC : UINT := 32384; (*Warning: The y coordinates of the node vector are not sorted in ascending or descending order.*)
  HCR_WARN_LIN_Y_NOT_ASC_DESC_S : UINT := 32385; (*Warning: Sorting of the y coordinates of the node vector is monotonic, but not strictly monotonic.*)
  HCR_WARN_PID_TF_TS : UINT := 32386; (*Warning: The filter time constant Tf of the differentiator is not larger than the corresponding task cycle time.*)
  HCR_WARN_PID_TN_NEG_TS : UINT := 32387; (*Warning:
PID: The integration time constant for I_Switch < 0 Tn_neg is not larger than the corresponding task cycle time.
Position controller: The integration time constant for movements in the 'negative' direction Tn_neg is not larger than the corresponding task cycle time.*)
  HCR_WARN_PID_TN_POS_TS : UINT := 32388; (*Warning:
PID: The integration time constant for I_Switch > 0 Tn_pos is not larger than the corresponding task cycle time.
Position controller: The integration time constant for movements in the 'positive' direction Tn_pos is not larger than the corresponding task cycle time.
Force controller: The integration time constant Tn entered is not larger than the corresponding task cycle time.*)
  HCR_WARN_PID_TV_TS : UINT := 32389; (*Warning: The differentiation time constant Tv of the differentiator is not larger than the corresponding task cycle time.*)
  HCR_WARN_PID_YADD_100 : UINT := 32390; (*Warning:
PID: The feed forward size Yadd was outside the permissible interval of [-100%, 100%] and has been limited accordingly.
Position controller: The feed forward speed v_add was outside the permissible interval of [-Internal.vCyl_sup, Internal.vCyl_sup] and has been limited accordingly.
Force controller: The feed forward volume flow Q_add was outside the permissible interval of [-Qnom_neg, Qnom_pos] and has been limited accordingly.*)
  HCR_WARN_PID_YI_MAX : UINT := 32391; (*Warning: The integrator's manipulated variable Yi has reached its maximum value.*)
  HCR_WARN_PID_YI_MIN : UINT := 32392; (*Warning: The integrator's manipulated variable Yi has reached its minimum value.*)
  HCR_WARN_PID_YMAN_MAX : UINT := 32393; (*Warning:
PID: The manipulated variable for manual operation Yman was set above the maximum permissible value Y_max and has been limited to this maximum.
Position controller: The speed of movement for manual operation v_man was set above the maximum permissible value v_max and has been limited to this maximum.
Force controller: The valve volume flow for manual operation Q_man was set above the maximum permissible value Q_max and has been limited to this maximum.*)
  HCR_WARN_PID_YMAN_MIN : UINT := 32394; (*Warning:
PID: The manipulated variable for manual operation Yman was set below the minimum permissible value Y_min and has been increased to this minimum.
Position controller: The speed of movement for manual operation v_man was set below the minimum permissible value v_min and has been increased to this minimum.
Force controller: The valve volume flow for manual operation Q_man was set below the minimum permissible value Q_min and has been increased to this minimum.*)
  HCR_WARN_PT12_T1_TS : UINT := 32395; (*Warning: The time constant T1 entered is not larger than the corresponding task cycle time.*)
  HCR_WARN_PT12_T1_ZERO : UINT := 32396; (*Warning: The time constant T1 = 0.*)
  HCR_WARN_PT12_T2_TS : UINT := 32397; (*Warning: The time constant T2 entered is not larger than the corresponding task cycle time.*)
  HCR_WARN_PT12_T2_ZERO : UINT := 32398; (*Warning: The time constant T2 = 0.*)
  HCR_WARN_PT1CP_T1_TS : UINT := 32399; (*Warning: The time constant T1 entered is not larger than the corresponding task cycle time.*)
  HCR_WARN_PT1CP_T1_ZERO : UINT := 32400; (*Warning: The time constant T1 = 0.*)
  HCR_WARN_PT2S_TF_TS : UINT := 32401; (*Warning: The filter time constant Tf entered is not larger than the corresponding task cycle time.*)
  HCR_WARN_SERVO_FF_CYL_NEG : UINT := 32402; (*Warning: Friction force in the 'negative' direction Ff_Cyl_neg < 0.*)
  HCR_WARN_SERVO_FF_CYL_POS : UINT := 32403; (*Warning: Friction force in the 'positive' direction Ff_Cyl_pos < 0.*)
  HCR_WARN_SERVO_P_CYL_NEG_HIGH : UINT := 32404; (*The calculated pressure for the 'negative' cylinder pressure chamber is too high.*)
  HCR_WARN_SERVO_P_CYL_NEG_LOW : UINT := 32405; (*Warning: The calculated pressure for the 'negative' cylinder pressure chamber is too low.*)
  HCR_WARN_SERVO_P_CYL_NEG_NEG : UINT := 32406; (*Warning: The measured or estimated pressure for the 'negative' cylinder pressure chamber is negative.*)
  HCR_WARN_SERVO_P_CYL_POS_HIGH : UINT := 32407; (*Warning: The calculated pressure for the 'positive' cylinder pressure chamber is too high.*)
  HCR_WARN_SERVO_P_CYL_POS_LOW : UINT := 32408; (*Warning: The calculated pressure for the 'positive' cylinder pressure chamber is too low.*)
  HCR_WARN_SERVO_P_CYL_POS_NEG : UINT := 32409; (*Warning: The measured or estimated pressure for the 'positive' cylinder pressure chamber is negative.*)
  HCR_WARN_SERVO_V_CYL_MAX : UINT := 32410; (*No longer used.*)
  HCR_WARN_SERVO_Y_MAX : UINT := 32411; (*Warning: The valve opening yValve has reached the maximum value (-1 or +1).*)
  HCR_WARN_SPF_MEM : UINT := 32412; (*Warning: An error occurred while allocating memory for the internal ring buffer.*)
  HCR_WARN_AUTOTUNE_KP_INVALID : UINT := 32413; (*No longer used.*)
  HCR_WARN_NOTCH_F0_FS : UINT := 32414; (*Warning: The filter frequency f0 is too high.*)
  HCR_WARN_IT1_T1_TS : UINT := 32416; (*Warning: The time constant T1 entered is not larger than the corresponding task cycle time.*)
  HCR_WARN_IT1_T1_ZERO : UINT := 32417; (*Warning: The time constant T1 = 0.*)
  HCR_WARN_IT1_TN_TS : UINT := 32418; (*Warning: The integration time constant Tn entered is not larger than the corresponding task cycle time.*)
  HCR_WARN_SFG_FP_END : UINT := 32419; (*Warning: Fp_end was selected equal to the value of the set force Fp_set when dFp_set ? 0.*)
  HCR_WARN_SFG_T_DELTA_ACT : UINT := 32420; (*Warning: The time t_delta_act, which was actually required for the profile generation, deviates massively from t_delta. However, a profile generation did occur.*)
  HCR_ERR_DISABLED : UINT := 65534; (*Error: The function block is disabled.*)
END_VAR
